FUNCTION_BLOCK FB_DomeState IMPLEMENTS I_DomeState

VAR
	TxBuffer	: ComBuffer;
	RxBuffer	: ComBuffer;
	pDome : POINTER TO FB_DomeControl;
END_VAR


METHOD CloseCommand : BOOL
LogIgnored(sCommand := 'close', sLevel := 'WARNING');
END_METHOD

METHOD FB_init : BOOL
VAR_INPUT
	bInitRetains : BOOL; // if TRUE, the retain variables are initialized (warm start / cold start)
	bInCopyCode : BOOL;  // if TRUE, the instance afterwards gets moved into the copy code (online change)
	pDome : POINTER TO FB_DomeControl;

END_VAR
THIS^.pDome := pDome;
END_METHOD


METHOD FoundError : BOOL
END_METHOD


METHOD HomeCommand : BOOL
LogIgnored(sCommand := 'home', sLevel := 'INFO');
END_METHOD

// #202: a line to the ADS log and to 50cm/Log (level WARNING or INFO)
METHOD LogEvent : BOOL
VAR_INPUT
	sText		: STRING(255);
	sLevel		: STRING(20) := 'INFO';
END_VAR
IF sLevel = 'WARNING' THEN
	ADSLOGSTR(ADSLOG_MSGTYPE_WARN OR ADSLOG_MSGTYPE_LOG, '%s', sText);
ELSE
	ADSLOGSTR(ADSLOG_MSGTYPE_HINT OR ADSLOG_MSGTYPE_LOG, '%s', sText);
END_IF
IF pDome <> 0 THEN
	IF pDome^.fbComm <> 0 THEN
		pDome^.fbComm.PublishLog(level := sLevel, message := sText);
	END_IF
END_IF
LogEvent := TRUE;
END_METHOD

// #202: a command that the state does not handle is dropped. Before, it was dropped without a trace: four dome_close
// went unnoticed while the dome was stuck in Closing.
METHOD LogIgnored : BOOL
VAR_INPUT
	sCommand	: STRING(20);
	sLevel		: STRING(20) := 'INFO';
END_VAR
LogIgnored := LogEvent(sText := CONCAT(CONCAT(CONCAT('Dome: ', sCommand), ' ignored in '), THIS^.StateID), sLevel := sLevel);
END_METHOD

METHOD MoveCommand : BOOL
END_METHOD


METHOD OpenCommand : BOOL
LogIgnored(sCommand := 'open', sLevel := 'INFO');
END_METHOD


METHOD ParkCommand : BOOL
LogIgnored(sCommand := 'park', sLevel := 'INFO');
END_METHOD


METHOD ResetCommand : BOOL
LogIgnored(sCommand := 'reset', sLevel := 'INFO');
END_METHOD

METHOD RunState : BOOL
VAR_INPUT
END_VAR
END_METHOD


PROPERTY StateID : STRING
GET
END_GET
END_PROPERTY


METHOD StopCommand : BOOL
LogIgnored(sCommand := 'stop', sLevel := 'INFO');
END_METHOD


METHOD SuccessfulFinished : BOOL
END_METHOD


METHOD TrackCommand : BOOL
END_METHOD

END_FUNCTION_BLOCK

(* stored: Version 1.1.0.1, ProductVersion 3.1.4024.15
   POU FB_DomeState: Id {ea26d2af-4995-4266-b54f-40ec64c0b456}, SpecialFunc None
   Method CloseCommand: Id {fb5de5a5-4a4d-45df-af61-071cca59aada}
   Method FB_init: Id {22775cbc-30f9-4d1f-bce5-a59c9bbf2750}
   Method FoundError: Id {42e4fbb5-dfee-4804-865e-273f0d90a6a6}
   Method HomeCommand: Id {573db44f-d9cf-4414-a9a5-4863a1da9bd1}
   Method LogEvent: Id {498ac7c6-4fe1-4a20-8711-0abc6d706da5}
   Method LogIgnored: Id {3f1c7a52-8d44-4b0e-9a6e-5b2f0c7d1e21}
   Method MoveCommand: Id {4d982227-1478-4c88-8c1e-b787654c2e0b}
   Method OpenCommand: Id {4d93018e-c4bd-4e1d-936d-acd45775b515}
   Method ParkCommand: Id {cf08df73-a434-4c35-812b-6a2a7fad3eb0}
   Method ResetCommand: Id {885bf905-2242-4d03-aaf3-a4eea3c12535}
   Method RunState: Id {551f815e-d0a0-47f3-a1bf-76df06e0e526}
   Property StateID: Id {33df2a26-65cb-4808-8c76-7a370a7d0a18}
   Get Get: Id {843679fd-fc2f-4f1a-b85a-a970f396d2f1}
   Method StopCommand: Id {b30e50be-4549-474b-9f4c-a5519dd17bc2}
   Method SuccessfulFinished: Id {062c433e-903b-4e33-8ead-c5a8ea2c9e66}
   Method TrackCommand: Id {dc19c696-fcda-492e-bd3e-af40a5f27b32} *)
